Staubli VAL3: stop.pgx

program stop()
// Stop motion and the IO task; preserve the actual gripper output.
begin
  // ============================================================
  // PARAR MOVIMIENTO Y EL ADAPTADOR, CONSERVANDO LA PINZA
  // ============================================================
  // Terminar primero la tarea de lectura de sensores.
  taskKill("physicalIO")
  resetMotion()
  ioReady = false
  cycleStep = -1

  // No llamar a open/close ni escribir valve1:
  // conservamos la salida real, sin soltar una posible pieza.
  // No retornar a jStart por una trayectoria pendiente de validar.
  // Un nuevo start comienza desde el principio; no es una reanudacion.
  putln("Stopped - gripper output unchanged; prepare cell before restart")
end
